// TIA Portal V21 export
DATA_BLOCK "IDB_AnaShared"   // DB14
// stored: InstanceOfName FB_AnaShared, InstanceOfType FB
"FB_AnaShared"
   // VAR_INPUT
   //    Pulse : Bool;
   // END_VAR
   // VAR_OUTPUT
   //    Count : Int;
   // END_VAR
   // VAR
   //    PulseEdge { S7_SetPoint := 'True'} : R_TRIG;
   // END_VAR
BEGIN
END_DATA_BLOCK
